(* Logix 5000 project; controller DSFW_Budzar vendor 1 type 14 code 154 rev 32.13; software revision 32.03; part 4 of 5 *)
(* tags used below, declared in another part *)
   PCV_Go_to_start_position_TMR : TIMER;
   Active_Setpoint : REAL;
   ALARMS : DINT[5];
   Batch_Mode_Enable : BOOL;
   C_101_AUX : ALIAS FOR Local:1:I.Data.8;
   Comp_1 : BudLib_Compressor;   // R507A Compressor 1
   Comp_1_Status : BOOL;
   Comp_404A_Timing_1 : BOOL;
   Comp_Start_Purge_Relay : BOOL;
   Compressor_R404A_Superheat : REAL;
   Compressor_Start_Request : BOOL;
   CR_109 : ALIAS FOR Local:1:O.Data.5;   // Compressor Motor Relay (Energizes Contactor C-101)
   EEV_101_Auto_Manual : BOOL;
   EEV_101_High_Range_CV_Max : REAL;
   EEV_101_High_Range_CV_Min : REAL;
   EEV_101_Low_Range_CV_Max : REAL;
   EEV_101_Low_Range_CV_Min : REAL;
   EEV_101_Manual_Percent : REAL;
   EEV_101_Mid_Range_CV_Max : REAL;
   EEV_101_Mid_Range_CV_Min : REAL;
   EEV_101_Pressure_Setpoint : REAL;
   EEV_101_Run_PIDE : BOOL;
   EEV_101_Run_Temp_PIDE : BOOL;
   EEV_101_Stop_PIDE : BOOL;
   EEV_101_Superheat_Setpoint : REAL;
   EEV_101_To_Purge : BOOL;   // Oil Management, Call For Purge with EEV-101
   EEV_102_Auto_Manual : BOOL;
   EEV_102_Manual_Percent : REAL;
   EEV_102_Run_PIDE : BOOL;
   EEV_102_Stop_PIDE : BOOL;
   EEV_102_Superheat_Setpoint : REAL;
   EEV_High_Range_Max_Temp : REAL;
   EEV_High_Range_Min_Temp : REAL;
   EEV_Low_Range_Max_Temp : REAL;
   EEV_Low_Range_Min_Temp : REAL;
   EEV_Manual_Relief_Delay : TIMER;   // Oil Management, Delay until Flush begins
   EEV_Manual_Relief_Timer : TIMER;   // Oil Management, Duration of Flush
   EEV_Mid_Range_Max_Temp : REAL;
   EEV_Mid_Range_Min_Temp : REAL;
   Engineering_Alarm_Reset : TIMER;
   Evaporator_R404A_Superheat : REAL;
   FIC_101_Run_PID : BOOL;
   High_Range_Max_Temp : REAL;
   High_Range_Min_Temp : REAL;
   HMI_EEV_101_CV : REAL;
   HMI_EEV_101_Lamp : BOOL;
   HMI_EEV_102_CV : REAL;
   HMI_EEV_102_Lamp : BOOL;
   HMI_Oil_Purge_Retries_Reset_Min : REAL;   // Oil Management, Compressor Runtime before resetting retry accumulator
   HMI_R404A_Hot_Gas_Switch_Delay : REAL;
   HMI_R404A_TCV_Toggle_SP : REAL;
   HMI_TCV_101_CV : REAL;
   HMI_TCV_101_Lamp : BOOL;
   HMI_TCV_102_CV : REAL;
   HMI_TCV_102_Lamp : BOOL;
   Low_Range_Max_Temp : REAL;
   Low_Range_Min_Temp : REAL;
   Mid_Range_Max_Temp : REAL;
   Mid_Range_Min_Temp : REAL;
   Oil_Purge_Fail : BOOL;   // Oil Management, This coil will energize after configured purge retries fail
   Oil_Purge_Relay : BOOL;   // Oil Management, Oil Purge Sequence Latch
   Oil_Purge_Retires_Enable : BOOL;
   Oil_Purge_Retries_ACC : DINT;   // Oil Management, Accumulated Oil Purges this low level
   Oil_Purge_Retries_Reset : TIMER;   // Oil Management, Reset Accumulator with 10-min without Low Level
   Oil_Purge_Retries_Reset1 : TIMER;   // Oil Management, Used to reset accuulated retries if compressor off.
   Oil_Purge_Retries_Reset_Remaining : REAL;   // Oil Management, Time remaining until reset retries accum
   Oil_Purge_Retries_SP : DINT;   // Oil Management, Desired Oil Purge Retries before Fault
   OMB_101 : ALIAS FOR Local:1:I.Data.12;
   ONS : DINT[3];   // One-Shots
   PCV_101_Flush_Limit : REAL;   // Temperature Limit (Deg F) to force Condenser Water Flush
   PCV_101_Flush_Time_Remaining : DINT;
   PCV_101_Flush_Timer : TIMER;   // PCV-101 Condenser Hot Water Flush Timer
   PCV_101_go_to_start_position : BOOL;
   PCV_101_Multiplexer : DINT;   // Selects controlling input to multiplxer
   PCV_101_Run_PIDE : BOOL;
   PCV_101_Stop_PIDE : BOOL;
   PT_104 : BL_Analog_Input;   // R404A Evaporator Suction Pressure
   PT_104_PID_Scale_Max : REAL;
   PT_104_PID_Scale_Min : REAL;
   Purge_Request : BOOL;   // Oil Management, Request to Purge
   R404A_HG_Switch_Delay : TIMER;
   R404A_HG_Switch_Off_Delay : TIMER;
   R404A_Hot_Gas_Toggle : BOOL;
   R404A_Hot_Gas_Toggle_Req : BOOL;
   R404A_OK_To_Run : BOOL;
   R404A_TCV_Toggle_SP_OFF : REAL;
   R404A_TCV_Toggle_SP_ON : REAL;
   R404A_TCV_Valve_Toggle : BOOL;
   REACTOR_BATCH_PID_START : BOOL;
   REACTOR_BATCH_PIDE_CV_AS_SP : REAL;
   Short_Cycle_1_Time_Remaining : DINT;
   System_Start : BOOL;   // System Start
   TCV_101_CV_RAW : ALIAS FOR Local:7:O.Ch3Data;   // TCV-101 Valve De-Scale Output (4000-20000)
   TCV_101_EVAP_PRESSURE_PIDE : PID_ENHANCED;   // TCV-101 Hot Gas Pressure PID loop
   TCV_101_EVAP_TEMPERATURE_PIDE : PID_ENHANCED;   // TCV-101 Evaporator Hot Gas Bypass PID loop
   TCV_101_High_Range_CV_Max : REAL;
   TCV_101_High_Range_CV_Min : REAL;
   TCV_101_Low_Range_CV_Max : REAL;
   TCV_101_Low_Range_CV_Min : REAL;
   TCV_101_Mid_Range_CV_Max : REAL;
   TCV_101_Mid_Range_CV_Min : REAL;
   TCV_101_Relay : BOOL;
   TCV_101_Run_PIDE : BOOL;
   TCV_101_Stop_PIDE : BOOL;
   TCV_102_CV_RAW : ALIAS FOR Local:8:O.Ch0Data;   // TCV-102 Valve De-Scale Output (4000-20000)
   TCV_102_Relay : BOOL;
   TCV_CV : REAL;   // TCV Loop Output Scaled (0-100%)
   TCV_Multiplexer : DINT;
   TCV_Mux : MULTIPLEXER;
   TE_101 : BL_Analog_Input;   // Process Supply Temperature
   TE_108 : BL_Analog_Input;   // CONDENSER CHILLED GLYCOL INLET TEMPERATURE SENSOR
   Valve_Flush_SP : REAL;
(* D_Refrigeration_Control, continued *)

ROUTINE Compressor_Control   (* ladder *)
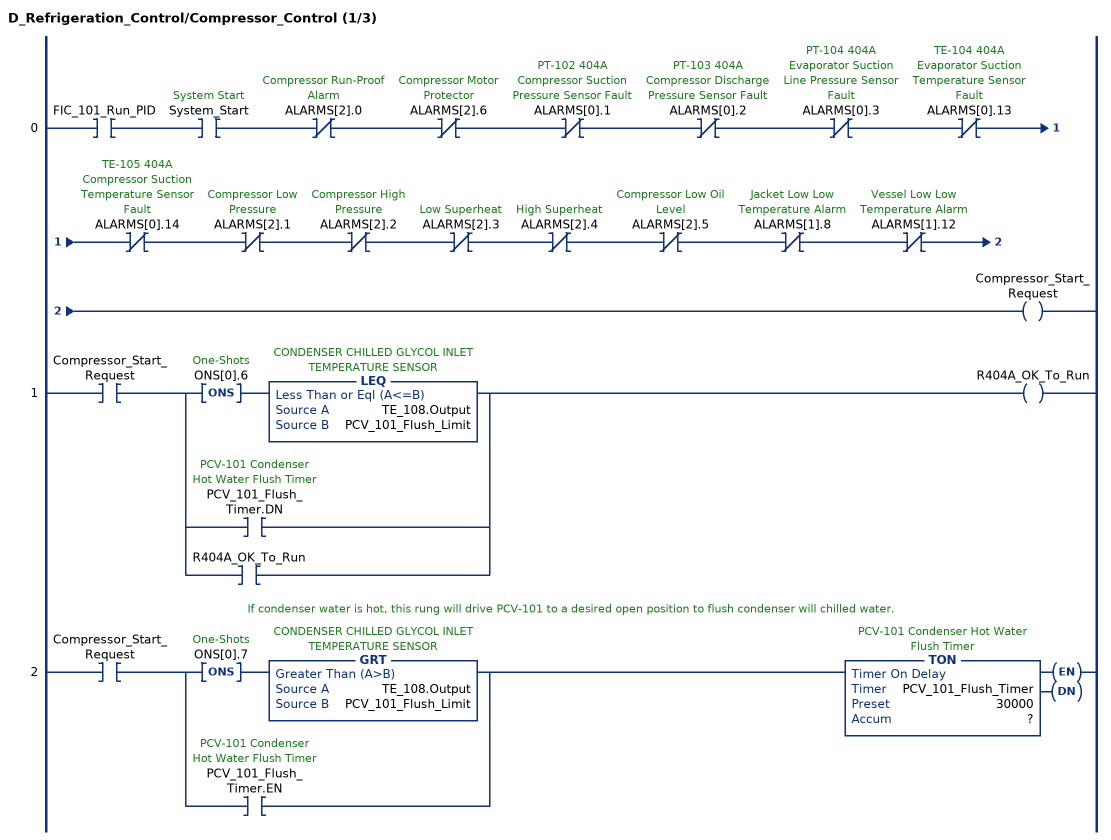
   0: XIC(FIC_101_Run_PID)XIC(System_Start)XIO(ALARMS[2].0)XIO(ALARMS[2].6)XIO(ALARMS[0].1)XIO(ALARMS[0].2)XIO(ALARMS[0].3)XIO(ALARMS[0].13)XIO(ALARMS[0].14)XIO(ALARMS[2].1)XIO(ALARMS[2].2)XIO(ALARMS[2].3)XIO(ALARMS[2].4)XIO(ALARMS[2].5)XIO(ALARMS[1].8)XIO(ALARMS[1].12)OTE(Compressor_Start_Request);
   1: XIC(Compressor_Start_Request)[ONS(ONS[0].6) LEQ(TE_108.Output,PCV_101_Flush_Limit) ,XIC(PCV_101_Flush_Timer.DN) ,XIC(R404A_OK_To_Run) ]OTE(R404A_OK_To_Run);
   // If condenser water is hot, this rung will drive PCV-101 to a desired open position to flush condenser will chilled water.
   2: XIC(Compressor_Start_Request)[ONS(ONS[0].7) GRT(TE_108.Output,PCV_101_Flush_Limit) ,XIC(PCV_101_Flush_Timer.EN) ]TON(PCV_101_Flush_Timer,?,?);
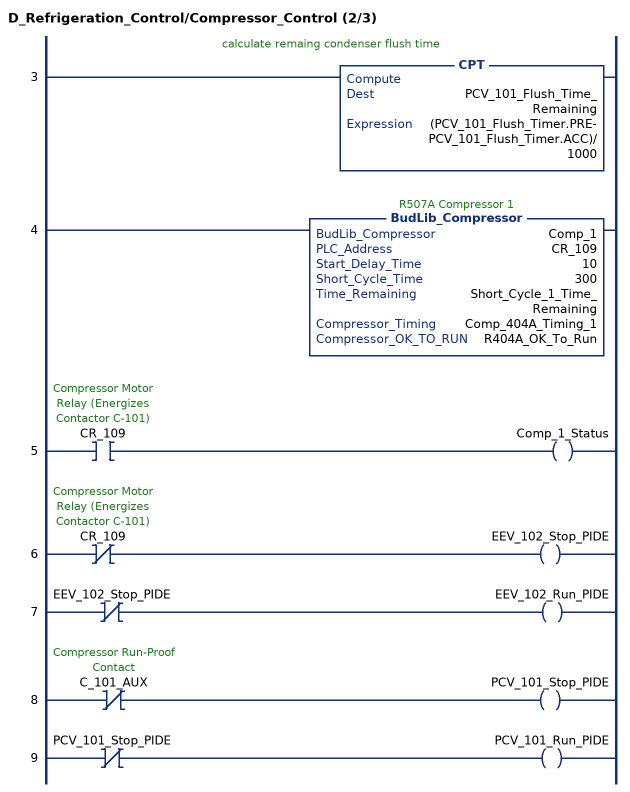
   // calculate remaing condenser flush time
   3: CPT(PCV_101_Flush_Time_Remaining,(PCV_101_Flush_Timer.PRE-PCV_101_Flush_Timer.ACC)/1000);
   4: BudLib_Compressor(Comp_1,CR_109,10,300,Short_Cycle_1_Time_Remaining,Comp_404A_Timing_1,R404A_OK_To_Run);
   5: XIC(CR_109)OTE(Comp_1_Status);
   6: XIO(CR_109)OTE(EEV_102_Stop_PIDE);
   7: XIO(EEV_102_Stop_PIDE)OTE(EEV_102_Run_PIDE);
   8: XIO(C_101_AUX)OTE(PCV_101_Stop_PIDE);
   9: XIO(PCV_101_Stop_PIDE)OTE(PCV_101_Run_PIDE);
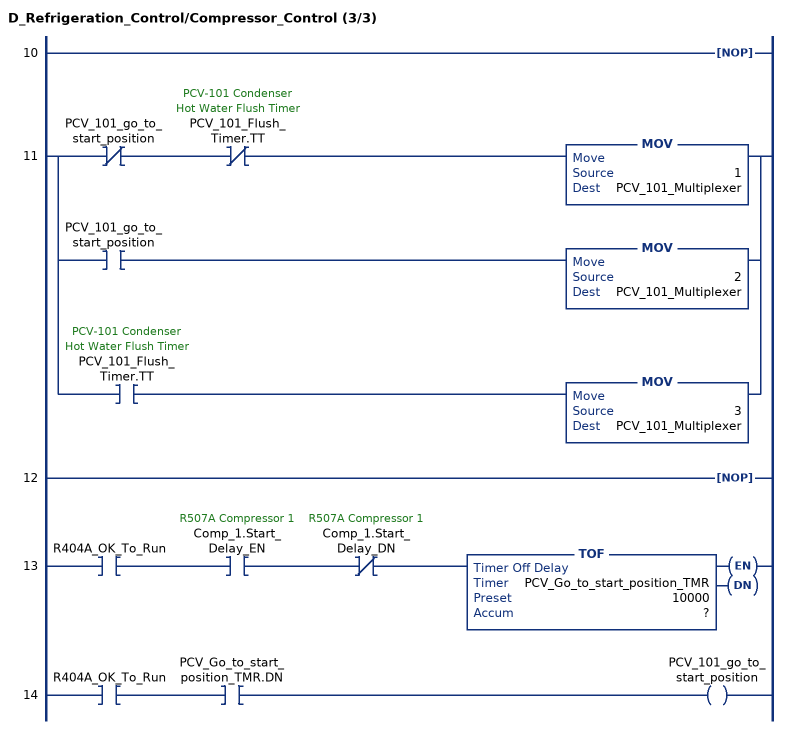
   10: NOP();
   11: [XIO(PCV_101_go_to_start_position) XIO(PCV_101_Flush_Timer.TT) MOV(1,PCV_101_Multiplexer) ,XIC(PCV_101_go_to_start_position) MOV(2,PCV_101_Multiplexer) ,XIC(PCV_101_Flush_Timer.TT) MOV(3,PCV_101_Multiplexer) ];
   12: NOP();
   13: XIC(R404A_OK_To_Run)XIC(Comp_1.Start_Delay_EN)XIO(Comp_1.Start_Delay_DN)TOF(PCV_Go_to_start_position_TMR,?,?);
   14: XIC(R404A_OK_To_Run)XIC(PCV_Go_to_start_position_TMR.DN)OTE(PCV_101_go_to_start_position);
END_ROUTINE

ROUTINE Evaporator_Control   (* ladder *)
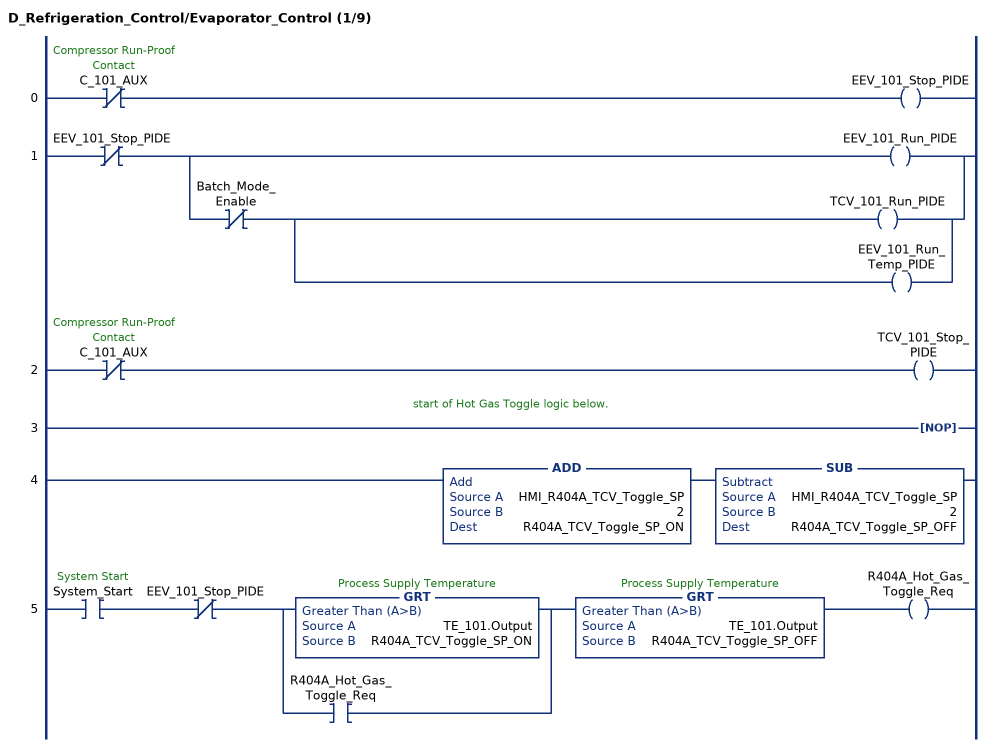
   0: XIO(C_101_AUX)OTE(EEV_101_Stop_PIDE);
   1: XIO(EEV_101_Stop_PIDE)[OTE(EEV_101_Run_PIDE) ,XIO(Batch_Mode_Enable) [OTE(TCV_101_Run_PIDE) ,OTE(EEV_101_Run_Temp_PIDE) ] ];
   2: XIO(C_101_AUX)OTE(TCV_101_Stop_PIDE);
   // start of Hot Gas Toggle logic below.
   3: NOP();
   4: ADD(HMI_R404A_TCV_Toggle_SP,2,R404A_TCV_Toggle_SP_ON)SUB(HMI_R404A_TCV_Toggle_SP,2,R404A_TCV_Toggle_SP_OFF);
   5: XIC(System_Start)XIO(EEV_101_Stop_PIDE)[GRT(TE_101.Output,R404A_TCV_Toggle_SP_ON) ,XIC(R404A_Hot_Gas_Toggle_Req) ]GRT(TE_101.Output,R404A_TCV_Toggle_SP_OFF)OTE(R404A_Hot_Gas_Toggle_Req);
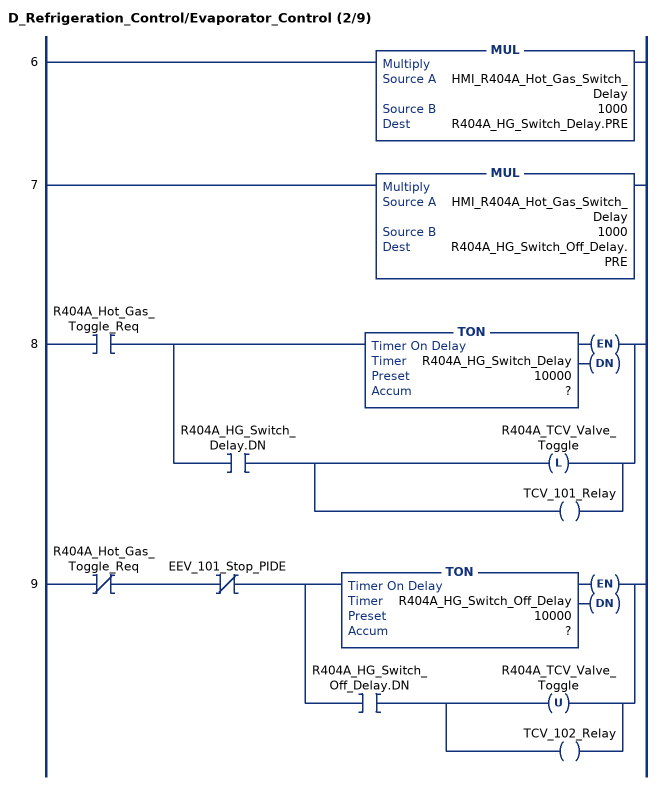
   6: MUL(HMI_R404A_Hot_Gas_Switch_Delay,1000,R404A_HG_Switch_Delay.PRE);
   7: MUL(HMI_R404A_Hot_Gas_Switch_Delay,1000,R404A_HG_Switch_Off_Delay.PRE);
   8: XIC(R404A_Hot_Gas_Toggle_Req)[TON(R404A_HG_Switch_Delay,?,?) ,XIC(R404A_HG_Switch_Delay.DN) [OTL(R404A_TCV_Valve_Toggle) ,OTE(TCV_101_Relay) ] ];
   9: XIO(R404A_Hot_Gas_Toggle_Req)XIO(EEV_101_Stop_PIDE)[TON(R404A_HG_Switch_Off_Delay,?,?) ,XIC(R404A_HG_Switch_Off_Delay.DN) [OTU(R404A_TCV_Valve_Toggle) ,OTE(TCV_102_Relay) ] ];
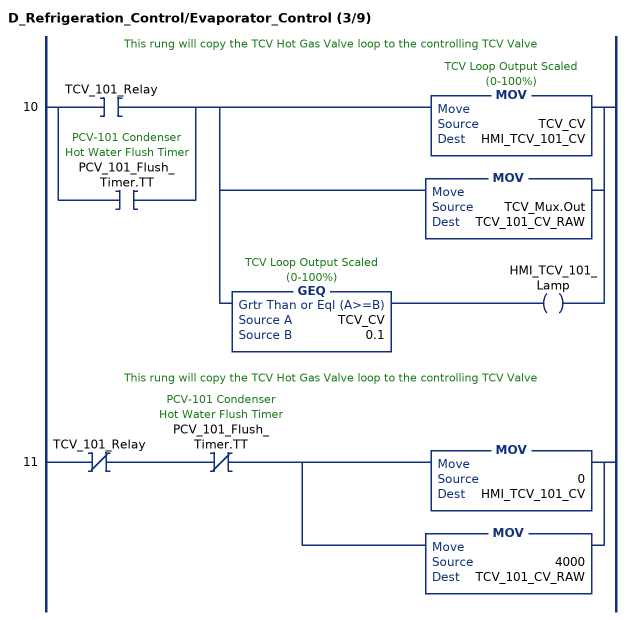
   // This rung will copy the TCV Hot Gas Valve loop to the controlling TCV Valve
   10: [XIC(TCV_101_Relay) ,XIC(PCV_101_Flush_Timer.TT) ][MOV(TCV_CV,HMI_TCV_101_CV) ,MOV(TCV_Mux.Out,TCV_101_CV_RAW) ,GEQ(TCV_CV,0.1) OTE(HMI_TCV_101_Lamp) ];
   // This rung will copy the TCV Hot Gas Valve loop to the controlling TCV Valve
   11: XIO(TCV_101_Relay)XIO(PCV_101_Flush_Timer.TT)[MOV(0,HMI_TCV_101_CV) ,MOV(4000,TCV_101_CV_RAW) ];
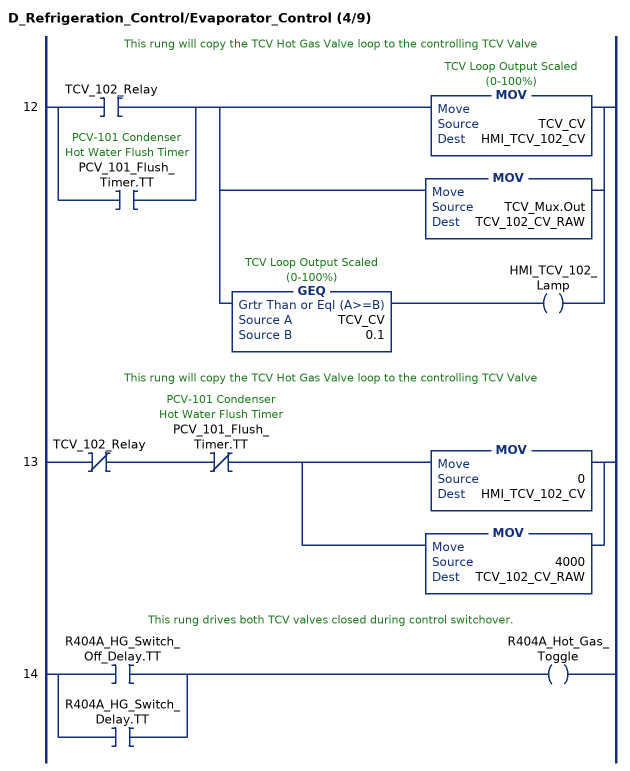
   // This rung will copy the TCV Hot Gas Valve loop to the controlling TCV Valve
   12: [XIC(TCV_102_Relay) ,XIC(PCV_101_Flush_Timer.TT) ][MOV(TCV_CV,HMI_TCV_102_CV) ,MOV(TCV_Mux.Out,TCV_102_CV_RAW) ,GEQ(TCV_CV,0.1) OTE(HMI_TCV_102_Lamp) ];
   // This rung will copy the TCV Hot Gas Valve loop to the controlling TCV Valve
   13: XIO(TCV_102_Relay)XIO(PCV_101_Flush_Timer.TT)[MOV(0,HMI_TCV_102_CV) ,MOV(4000,TCV_102_CV_RAW) ];
   // This rung drives both TCV valves closed during control switchover.
   14: [XIC(R404A_HG_Switch_Off_Delay.TT) ,XIC(R404A_HG_Switch_Delay.TT) ]OTE(R404A_Hot_Gas_Toggle);
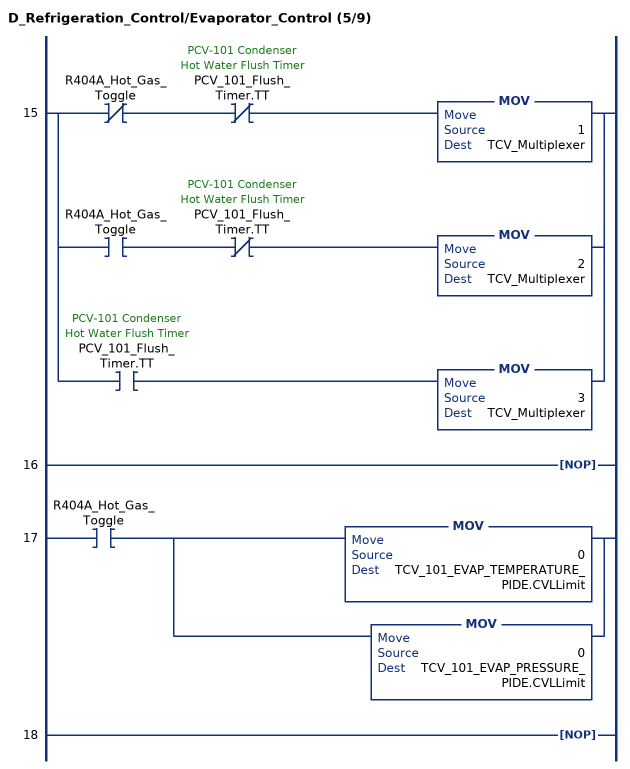
   15: [XIO(R404A_Hot_Gas_Toggle) XIO(PCV_101_Flush_Timer.TT) MOV(1,TCV_Multiplexer) ,XIC(R404A_Hot_Gas_Toggle) XIO(PCV_101_Flush_Timer.TT) MOV(2,TCV_Multiplexer) ,XIC(PCV_101_Flush_Timer.TT) MOV(3,TCV_Multiplexer) ];
   16: NOP();
   17: XIC(R404A_Hot_Gas_Toggle)[MOV(0,TCV_101_EVAP_TEMPERATURE_PIDE.CVLLimit) ,MOV(0,TCV_101_EVAP_PRESSURE_PIDE.CVLLimit) ];
   18: NOP();
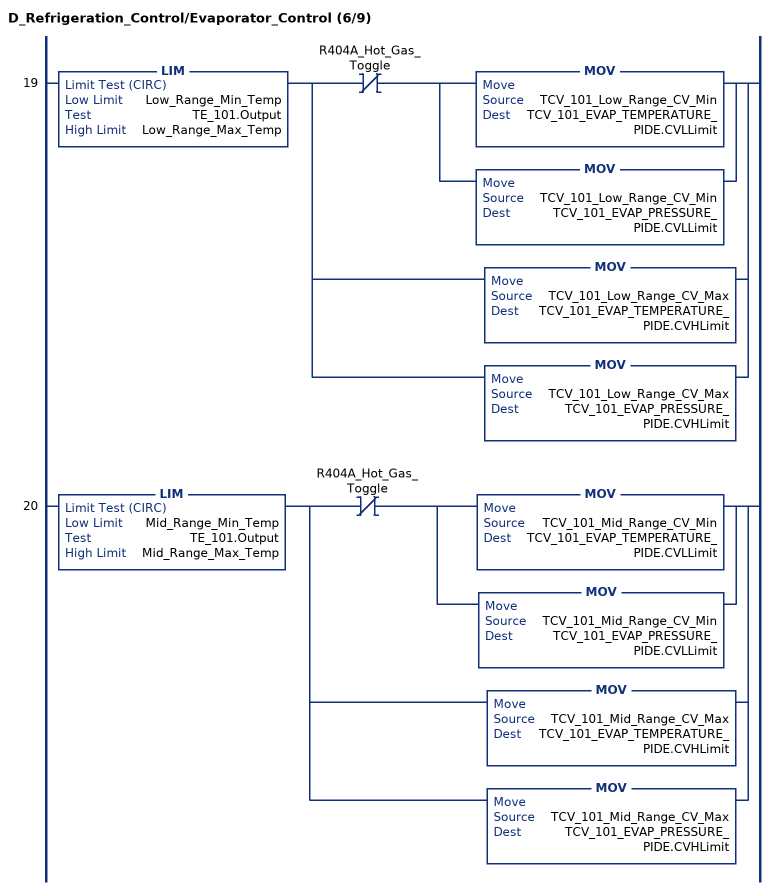
   19: LIM(Low_Range_Min_Temp,TE_101.Output,Low_Range_Max_Temp)[XIO(R404A_Hot_Gas_Toggle) [MOV(TCV_101_Low_Range_CV_Min,TCV_101_EVAP_TEMPERATURE_PIDE.CVLLimit) ,MOV(TCV_101_Low_Range_CV_Min,TCV_101_EVAP_PRESSURE_PIDE.CVLLimit) ] ,[MOV(TCV_101_Low_Range_CV_Max,TCV_101_EVAP_TEMPERATURE_PIDE.CVHLimit) ,MOV(TCV_101_Low_Range_CV_Max,TCV_101_EVAP_PRESSURE_PIDE.CVHLimit) ] ];
   20: LIM(Mid_Range_Min_Temp,TE_101.Output,Mid_Range_Max_Temp)[XIO(R404A_Hot_Gas_Toggle) [MOV(TCV_101_Mid_Range_CV_Min,TCV_101_EVAP_TEMPERATURE_PIDE.CVLLimit) ,MOV(TCV_101_Mid_Range_CV_Min,TCV_101_EVAP_PRESSURE_PIDE.CVLLimit) ] ,[MOV(TCV_101_Mid_Range_CV_Max,TCV_101_EVAP_TEMPERATURE_PIDE.CVHLimit) ,MOV(TCV_101_Mid_Range_CV_Max,TCV_101_EVAP_PRESSURE_PIDE.CVHLimit) ] ];
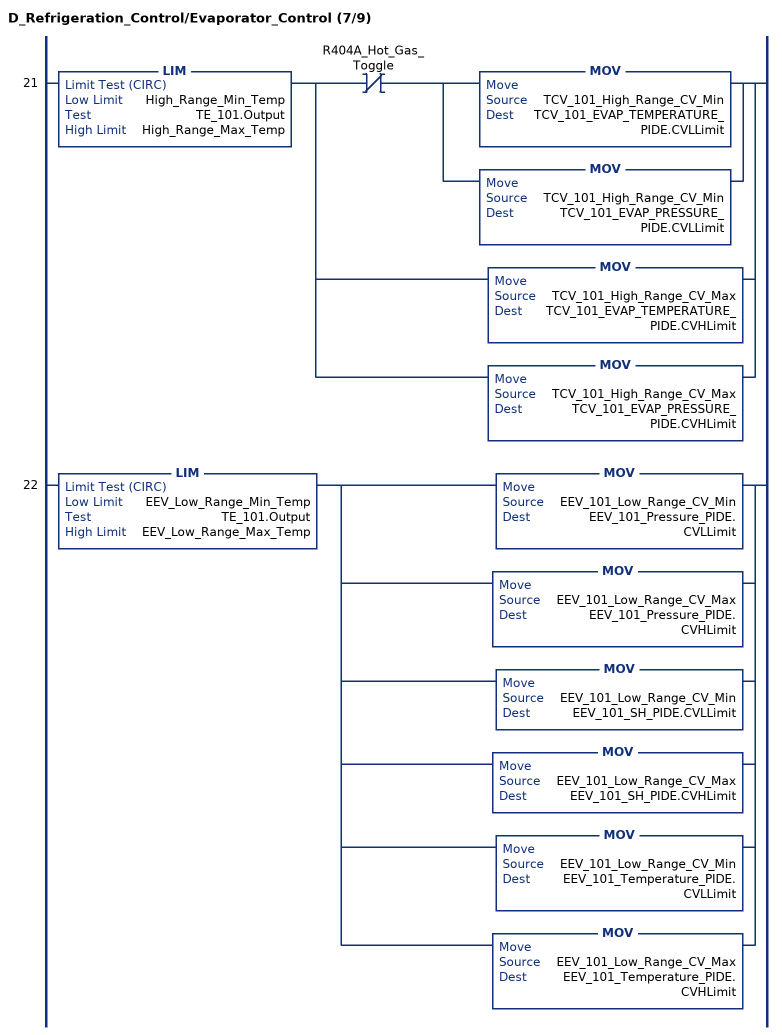
   21: LIM(High_Range_Min_Temp,TE_101.Output,High_Range_Max_Temp)[XIO(R404A_Hot_Gas_Toggle) [MOV(TCV_101_High_Range_CV_Min,TCV_101_EVAP_TEMPERATURE_PIDE.CVLLimit) ,MOV(TCV_101_High_Range_CV_Min,TCV_101_EVAP_PRESSURE_PIDE.CVLLimit) ] ,[MOV(TCV_101_High_Range_CV_Max,TCV_101_EVAP_TEMPERATURE_PIDE.CVHLimit) ,MOV(TCV_101_High_Range_CV_Max,TCV_101_EVAP_PRESSURE_PIDE.CVHLimit) ] ];
   22: LIM(EEV_Low_Range_Min_Temp,TE_101.Output,EEV_Low_Range_Max_Temp)[MOV(EEV_101_Low_Range_CV_Min,EEV_101_Pressure_PIDE.CVLLimit) ,MOV(EEV_101_Low_Range_CV_Max,EEV_101_Pressure_PIDE.CVHLimit) ,MOV(EEV_101_Low_Range_CV_Min,EEV_101_SH_PIDE.CVLLimit) ,MOV(EEV_101_Low_Range_CV_Max,EEV_101_SH_PIDE.CVHLimit) ,MOV(EEV_101_Low_Range_CV_Min,EEV_101_Temperature_PIDE.CVLLimit) ,MOV(EEV_101_Low_Range_CV_Max,EEV_101_Temperature_PIDE.CVHLimit) ];
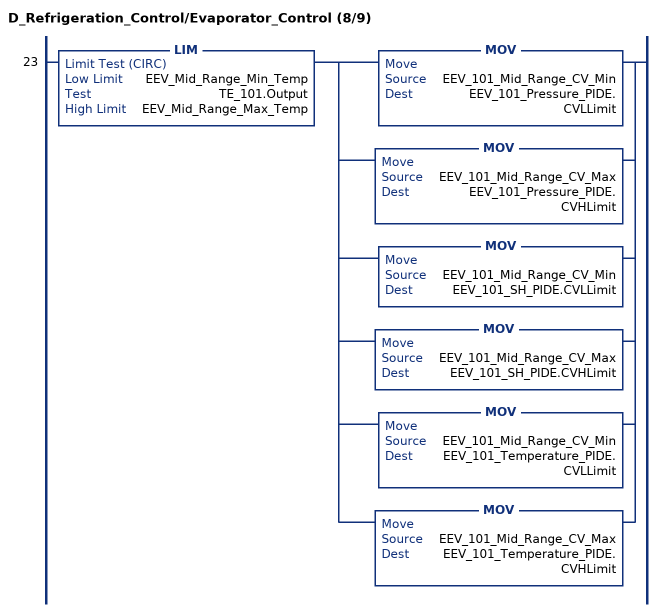
   23: LIM(EEV_Mid_Range_Min_Temp,TE_101.Output,EEV_Mid_Range_Max_Temp)[MOV(EEV_101_Mid_Range_CV_Min,EEV_101_Pressure_PIDE.CVLLimit) ,MOV(EEV_101_Mid_Range_CV_Max,EEV_101_Pressure_PIDE.CVHLimit) ,MOV(EEV_101_Mid_Range_CV_Min,EEV_101_SH_PIDE.CVLLimit) ,MOV(EEV_101_Mid_Range_CV_Max,EEV_101_SH_PIDE.CVHLimit) ,MOV(EEV_101_Mid_Range_CV_Min,EEV_101_Temperature_PIDE.CVLLimit) ,MOV(EEV_101_Mid_Range_CV_Max,EEV_101_Temperature_PIDE.CVHLimit) ];
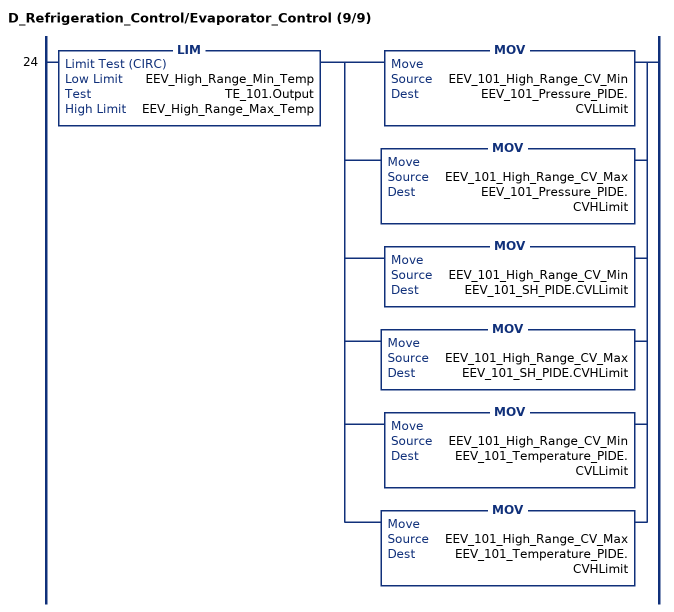
   24: LIM(EEV_High_Range_Min_Temp,TE_101.Output,EEV_High_Range_Max_Temp)[MOV(EEV_101_High_Range_CV_Min,EEV_101_Pressure_PIDE.CVLLimit) ,MOV(EEV_101_High_Range_CV_Max,EEV_101_Pressure_PIDE.CVHLimit) ,MOV(EEV_101_High_Range_CV_Min,EEV_101_SH_PIDE.CVLLimit) ,MOV(EEV_101_High_Range_CV_Max,EEV_101_SH_PIDE.CVHLimit) ,MOV(EEV_101_High_Range_CV_Min,EEV_101_Temperature_PIDE.CVLLimit) ,MOV(EEV_101_High_Range_CV_Max,EEV_101_Temperature_PIDE.CVHLimit) ];
END_ROUTINE

ROUTINE Oil_Management   (* ladder *)
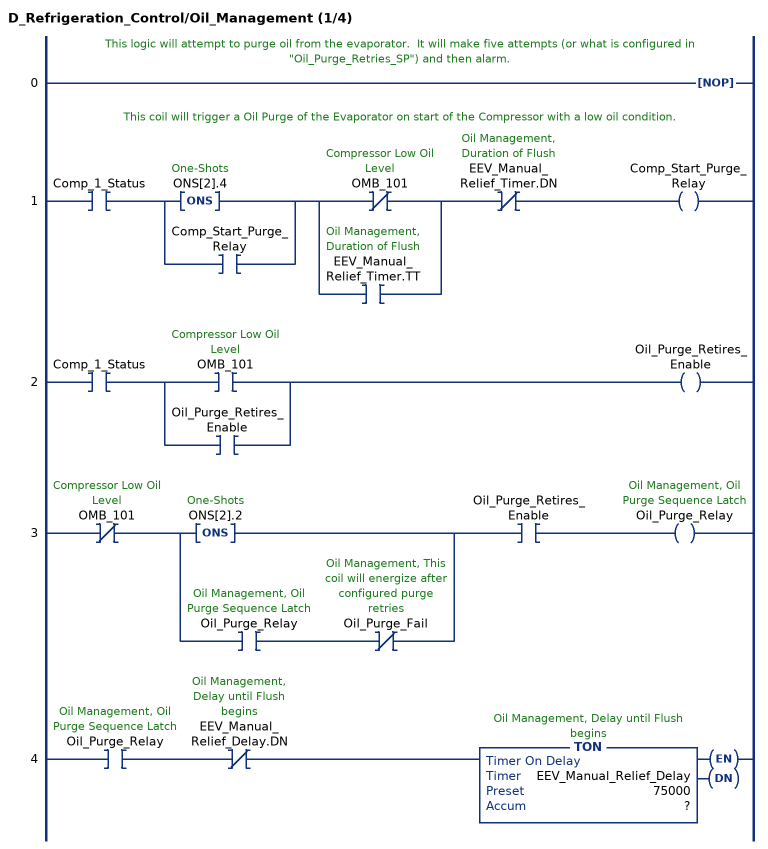
   // This logic will attempt to purge oil from the evaporator.  It will make five attempts (or what is configured in "Oil_Purge_Retries_SP") and then alarm.
   0: NOP();
   // This coil will trigger a Oil Purge of the Evaporator on start of the Compressor with a low oil condition.
   1: XIC(Comp_1_Status)[ONS(ONS[2].4) ,XIC(Comp_Start_Purge_Relay) ][XIO(OMB_101) ,XIC(EEV_Manual_Relief_Timer.TT) ]XIO(EEV_Manual_Relief_Timer.DN)OTE(Comp_Start_Purge_Relay);
   2: XIC(Comp_1_Status)[XIC(OMB_101) ,XIC(Oil_Purge_Retires_Enable) ]OTE(Oil_Purge_Retires_Enable);
   3: XIO(OMB_101)[ONS(ONS[2].2) ,XIC(Oil_Purge_Relay) XIO(Oil_Purge_Fail) ]XIC(Oil_Purge_Retires_Enable)OTE(Oil_Purge_Relay);
   4: XIC(Oil_Purge_Relay)XIO(EEV_Manual_Relief_Delay.DN)TON(EEV_Manual_Relief_Delay,?,?);
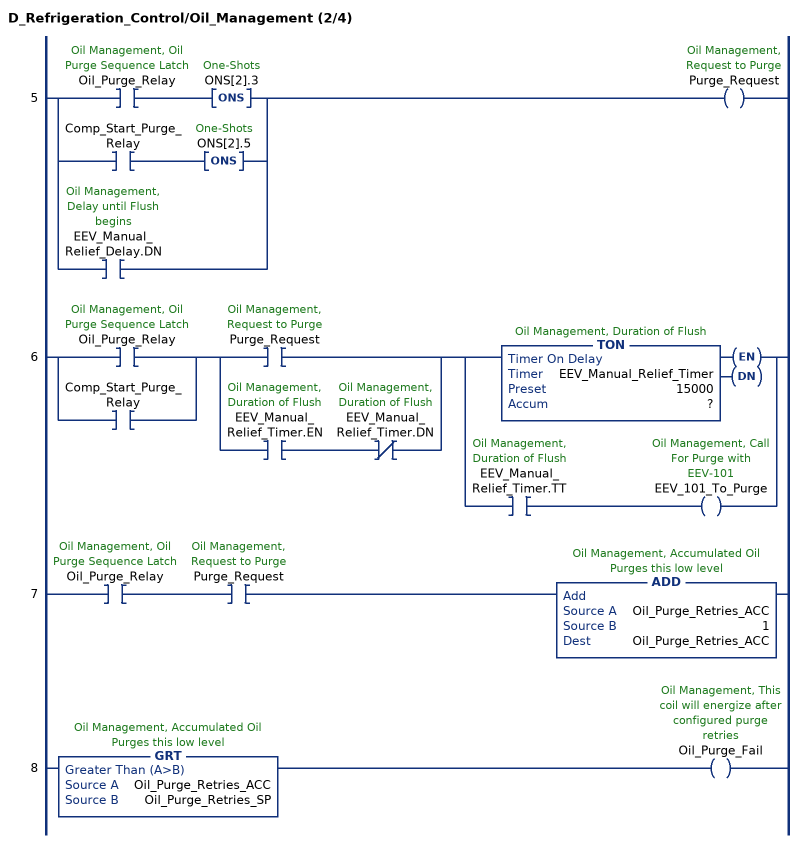
   5: [XIC(Oil_Purge_Relay) ONS(ONS[2].3) ,XIC(Comp_Start_Purge_Relay) ONS(ONS[2].5) ,XIC(EEV_Manual_Relief_Delay.DN) ]OTE(Purge_Request);
   6: [XIC(Oil_Purge_Relay) ,XIC(Comp_Start_Purge_Relay) ][XIC(Purge_Request) ,XIC(EEV_Manual_Relief_Timer.EN) XIO(EEV_Manual_Relief_Timer.DN) ][TON(EEV_Manual_Relief_Timer,?,?) ,XIC(EEV_Manual_Relief_Timer.TT) OTE(EEV_101_To_Purge) ];
   7: XIC(Oil_Purge_Relay)XIC(Purge_Request)ADD(Oil_Purge_Retries_ACC,1,Oil_Purge_Retries_ACC);
   8: GRT(Oil_Purge_Retries_ACC,Oil_Purge_Retries_SP)OTE(Oil_Purge_Fail);
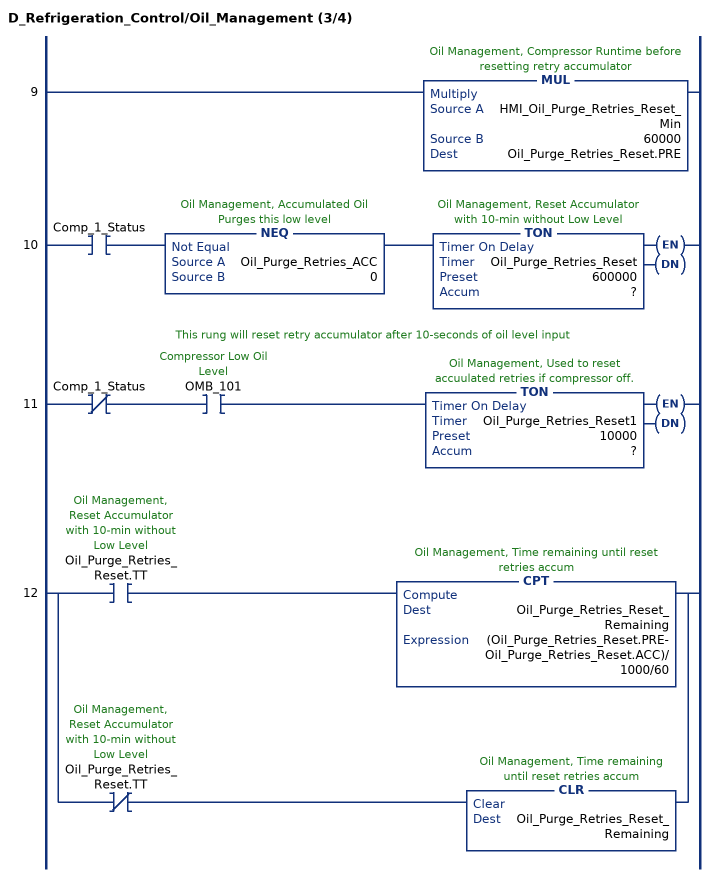
   9: MUL(HMI_Oil_Purge_Retries_Reset_Min,60000,Oil_Purge_Retries_Reset.PRE);
   10: XIC(Comp_1_Status)NEQ(Oil_Purge_Retries_ACC,0)TON(Oil_Purge_Retries_Reset,?,?);
   // This rung will reset retry accumulator after 10-seconds of oil level input
   11: XIO(Comp_1_Status)XIC(OMB_101)TON(Oil_Purge_Retries_Reset1,?,?);
   12: [XIC(Oil_Purge_Retries_Reset.TT) CPT(Oil_Purge_Retries_Reset_Remaining,(Oil_Purge_Retries_Reset.PRE-Oil_Purge_Retries_Reset.ACC)/1000/60) ,XIO(Oil_Purge_Retries_Reset.TT) CLR(Oil_Purge_Retries_Reset_Remaining) ];
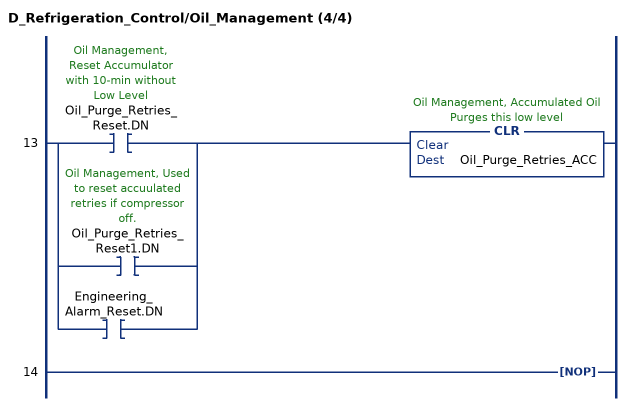
   13: [XIC(Oil_Purge_Retries_Reset.DN) ,XIC(Oil_Purge_Retries_Reset1.DN) ,XIC(Engineering_Alarm_Reset.DN) ]CLR(Oil_Purge_Retries_ACC);
   14: NOP();
END_ROUTINE

ROUTINE Routine_Schedule   (* ladder *)
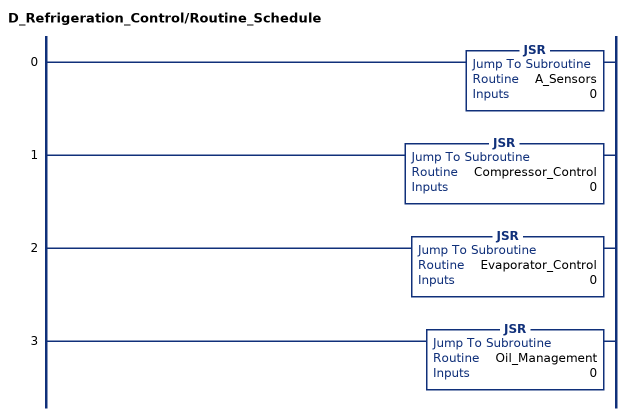
   0: JSR(A_Sensors,0);
   1: JSR(Compressor_Control,0);
   2: JSR(Evaporator_Control,0);
   3: JSR(Oil_Management,0);
END_ROUTINE
END_PROGRAM

PROGRAM EEV_PID   (* main routine Routine_Schedule *)
VAR
   BOR_01 : FBD_BOOLEAN_OR;
   BOR_02 : FBD_BOOLEAN_OR;
   ESEL_01 : SELECT_ENHANCED := (In1 := 4000.0, In2 := 4000.0, In3 := 4000.0, InsUsed := 3, SelectorMode := 2, OperSelector := 1, ProgProgReq := 1, Out := 4000.0, SelectedIn := 1, ProgOper := 1);
   ESEL_02 : SELECT_ENHANCED := (In1 := 4000.0, In2 := 4000.0, In3 := 4000.0, InsUsed := 3, SelectorMode := 2, OperSelector := 1, ProgProgReq := 1, Out := 4000.0, SelectedIn := 1, ProgOper := 1);
   ESEL_03 : SELECT_ENHANCED := (In1 := 6400.0, In2 := 12000.0, In3 := 12000.0, InsUsed := 3, SelectorMode := 2, OperSelector := 1, Out := 6400.0, SelectedIn := 1, ProgOper := 1);
   GEQ_01 : FBD_COMPARE := (SourceA := 4000.0, SourceB := 4100.0);
   GEQ_02 : FBD_COMPARE := (SourceB := 0.5);
   GEQ_03 : FBD_COMPARE := (SourceA := 4000.0, SourceB := 4100.0);
   GEQ_04 : FBD_COMPARE := (SourceA := 4000.0, SourceB := 4100.0);
   GEQ_05 : FBD_COMPARE := (SourceB := 0.5);
   GEQ_06 : FBD_COMPARE := (SourceA := 6400.0, SourceB := 4100.0, Dest := 1);
   MUX_01 : MULTIPLEXER := (In1 := 4000.0, In2 := 10400.0, Selector := 1, Out := 4000.0);
   PIDE_01 : PID_ENHANCED := (PVEUMax := 140.0, SPProg := 20.0, SPHLimit := 125.0, RatioProg := 1.0, RatioOper := 1.0, RatioHLimit := 1.0, RatioLLimit := 1.0, CVEUMax := 100.0, CVHLimit := 100.0, ControlAction := 1, PGain := 2.0, IGain := 1.0, PVEDerivative := 1, DSmoothing := 1, PVTracking := 1, ProgOverrideReq := 1, RTSTime := 1, InitPrimary := 1, Ratio := 1.0, Override := 1, DeltaT := 0.1);
   PIDE_02 : PID_ENHANCED := (PVEUMax := 140.0, SPProg := 20.0, SPHLimit := 125.0, RatioProg := 1.0, RatioOper := 1.0, RatioHLimit := 1.0, RatioLLimit := 1.0, CVEUMax := 100.0, CVHLimit := 100.0, ControlAction := 1, PGain := 2.0, IGain := 1.0, PVEDerivative := 1, DSmoothing := 1, PVTracking := 1, ProgOverrideReq := 1, RTSTime := 1, InitPrimary := 1, Ratio := 1.0, Override := 1, DeltaT := 0.1);
   PIDE_03 : PID_ENHANCED := (PVEUMax := 140.0, SPProg := 20.0, SPHLimit := 125.0, RatioProg := 1.0, RatioOper := 1.0, RatioHLimit := 1.0, RatioLLimit := 1.0, CVEUMax := 100.0, CVHLimit := 100.0, ControlAction := 1, PGain := 2.0, IGain := 1.0, PVEDerivative := 1, DSmoothing := 1, PVTracking := 1, ProgOverrideReq := 1, RTSTime := 1, InitPrimary := 1, Ratio := 1.0, Override := 1, DeltaT := 0.1);
   SCL_01 : SCALE := (In := 35.0, InRawMax := 60.0, InEUMax := 20000.0, InEUMin := 4000.0, Out := 13333.334);
   SCL_02 : SCALE := (In := 4000.0, InRawMax := 20000.0, InRawMin := 4000.0, InEUMax := 100.0);
   SCL_03 : SCALE := (In := 4000.0, InRawMax := 20000.0, InRawMin := 4000.0, InEUMax := 100.0);
   SCL_04 : SCALE := (In := 6400.0, InRawMax := 20000.0, InRawMin := 4000.0, InEUMax := 100.0, Out := 15.0);
   SCL_05 : SCALE := (In := 4000.0, InRawMax := 20000.0, InRawMin := 4000.0, InEUMax := 100.0);
   SEL_01 : SELECT := (In1 := 4000.0, In2 := 13600.0, Out := 4000.0);
END_VAR

ROUTINE R404A_EEV_PIDS   (* function block diagram *)
   SHEET 1
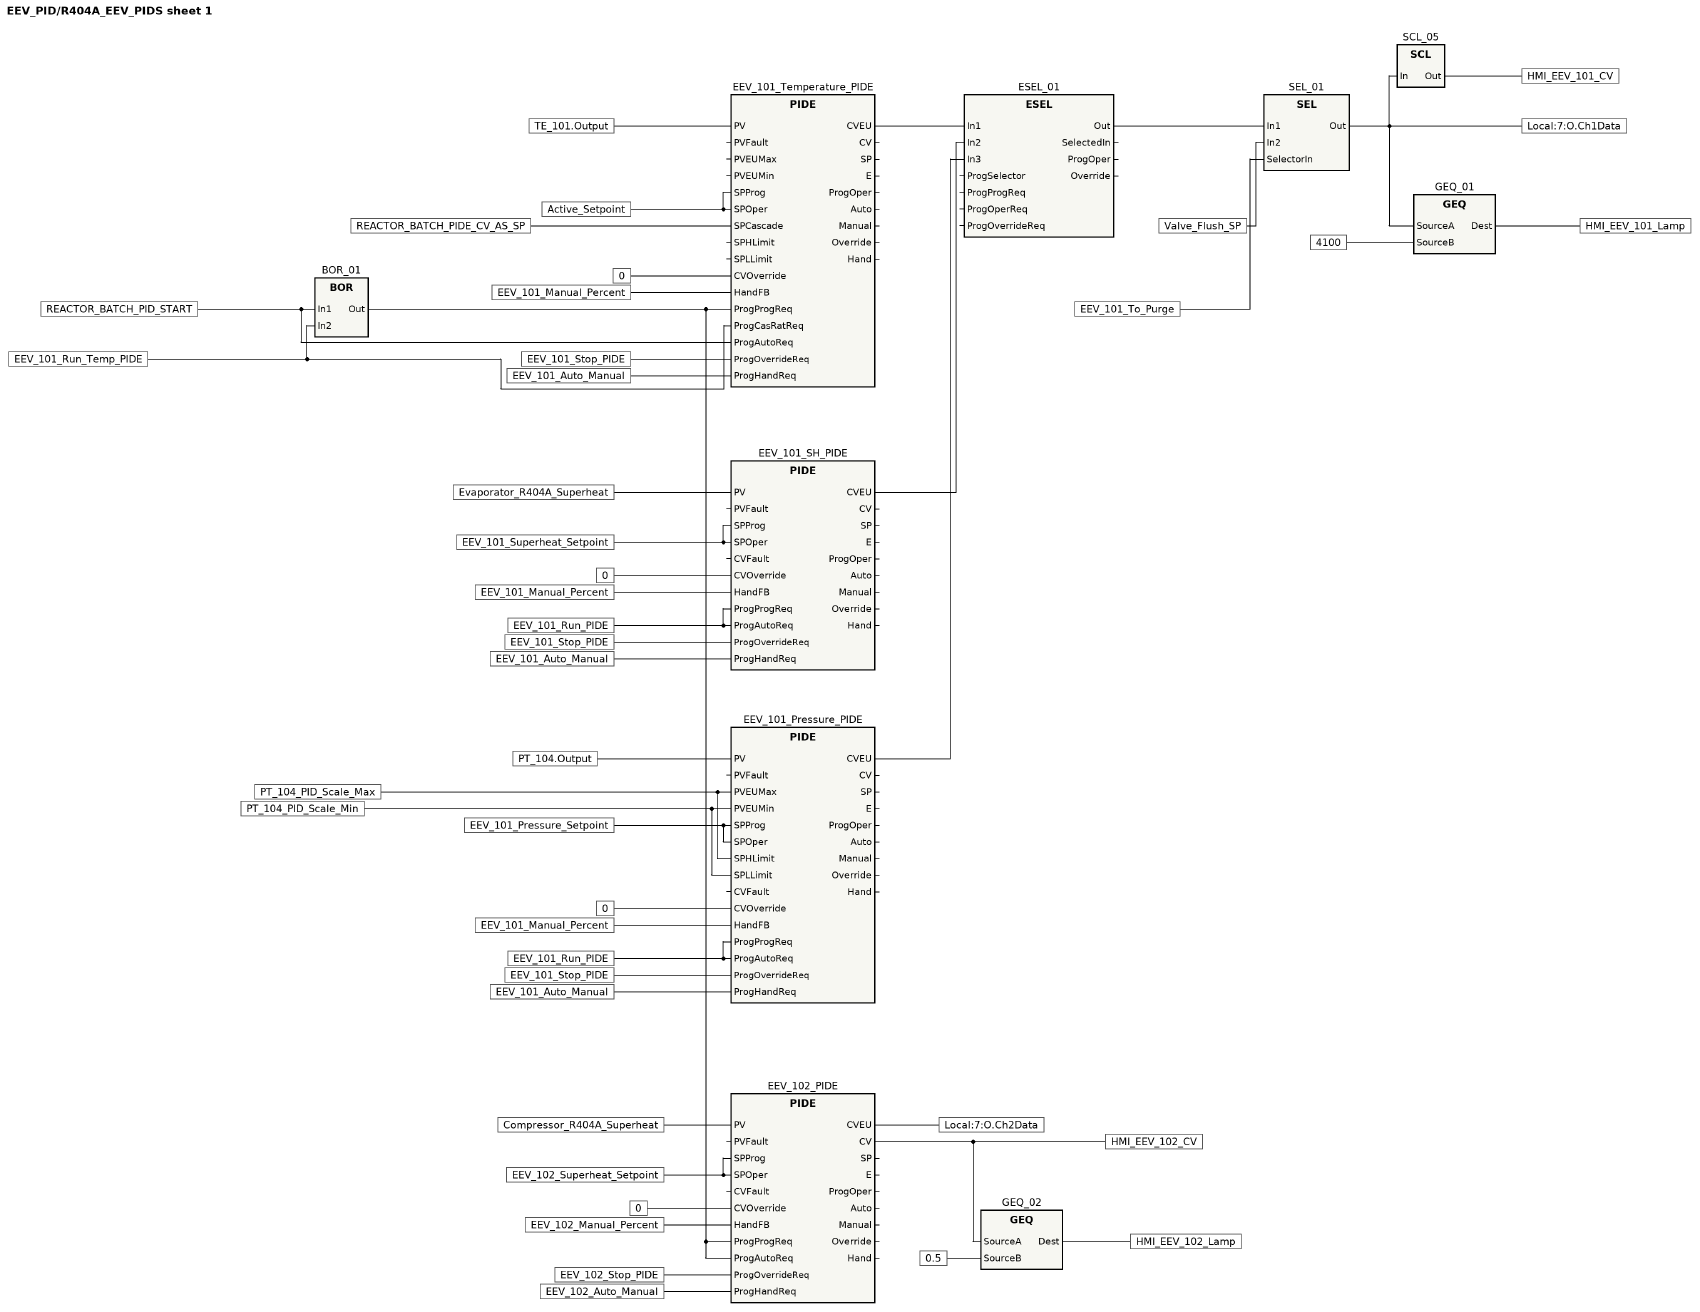
   BOR_01 : BOR(In1 := REACTOR_BATCH_PID_START, In2 := EEV_101_Run_Temp_PIDE);
   EEV_101_Temperature_PIDE : PIDE(PV := TE_101.Output, SPProg := Active_Setpoint, SPOper := Active_Setpoint, SPCascade := REACTOR_BATCH_PIDE_CV_AS_SP, CVOverride := 0, HandFB := EEV_101_Manual_Percent, ProgProgReq := BOR_01.Out, ProgCasRatReq := REACTOR_BATCH_PID_START, ProgAutoReq := EEV_101_Run_Temp_PIDE, ProgOverrideReq := EEV_101_Stop_PIDE, ProgHandReq := EEV_101_Auto_Manual);   // unwired pins: PVFault PVEUMax PVEUMin SPHLimit SPLLimit CV SP E ProgOper Auto Manual Override Hand
   EEV_101_SH_PIDE : PIDE(PV := Evaporator_R404A_Superheat, SPProg := EEV_101_Superheat_Setpoint, SPOper := EEV_101_Superheat_Setpoint, CVOverride := 0, HandFB := EEV_101_Manual_Percent, ProgProgReq := EEV_101_Run_PIDE, ProgAutoReq := EEV_101_Run_PIDE, ProgOverrideReq := EEV_101_Stop_PIDE, ProgHandReq := EEV_101_Auto_Manual);   // unwired pins: PVFault CVFault CV SP E ProgOper Auto Manual Override Hand
   EEV_101_Pressure_PIDE : PIDE(PV := PT_104.Output, PVEUMax := PT_104_PID_Scale_Max, PVEUMin := PT_104_PID_Scale_Min, SPProg := EEV_101_Pressure_Setpoint, SPOper := EEV_101_Pressure_Setpoint, SPHLimit := PT_104_PID_Scale_Max, SPLLimit := PT_104_PID_Scale_Min, CVOverride := 0, HandFB := EEV_101_Manual_Percent, ProgProgReq := EEV_101_Run_PIDE, ProgAutoReq := EEV_101_Run_PIDE, ProgOverrideReq := EEV_101_Stop_PIDE, ProgHandReq := EEV_101_Auto_Manual);   // unwired pins: PVFault CVFault CV SP E ProgOper Auto Manual Override Hand
   EEV_102_PIDE : PIDE(PV := Compressor_R404A_Superheat, SPProg := EEV_102_Superheat_Setpoint, SPOper := EEV_102_Superheat_Setpoint, CVOverride := 0, HandFB := EEV_102_Manual_Percent, ProgProgReq := BOR_01.Out, ProgAutoReq := BOR_01.Out, ProgOverrideReq := EEV_102_Stop_PIDE, ProgHandReq := EEV_102_Auto_Manual);   // unwired pins: PVFault CVFault SP E ProgOper Auto Manual Override Hand
   Local:7:O.Ch2Data := EEV_102_PIDE.CVEU;
   ESEL_01 : ESEL(In1 := EEV_101_Temperature_PIDE.CVEU, In2 := EEV_101_SH_PIDE.CVEU, In3 := EEV_101_Pressure_PIDE.CVEU);   // unwired pins: ProgSelector ProgProgReq ProgOperReq ProgOverrideReq SelectedIn ProgOper Override
   GEQ_02 : GEQ(SourceA := EEV_102_PIDE.CV, SourceB := 0.5);
   HMI_EEV_102_CV := EEV_102_PIDE.CV;
   HMI_EEV_102_Lamp := GEQ_02.Dest;
   SEL_01 : SEL(In1 := ESEL_01.Out, In2 := Valve_Flush_SP, SelectorIn := EEV_101_To_Purge);
   SCL_05 : SCL(In := SEL_01.Out);
   GEQ_01 : GEQ(SourceA := SEL_01.Out, SourceB := 4100);
   HMI_EEV_101_CV := SCL_05.Out;
   Local:7:O.Ch1Data := SEL_01.Out;
   HMI_EEV_101_Lamp := GEQ_01.Dest;
END_ROUTINE
